(* IEC 61131-3 sources: iolistgen/tests_support/pl_stub/src/DUTs/Common, 7 files *)

(* ---- E_CmdResult.dut.st ---- *)
// Назначение: заглушка plc-process-lib 1.0.0 для проверки типов сгенерированного кода без CODESYS
//             (API.md, раздел 4.1); не библиотека — тел и внутренних переменных нет
// Автор:      kr0nsch
// Версия:     1.0.0 (выпуск библиотеки)
// Документ:   docs/GENERATORS.md, раздел «Проверка ST без CODESYS»
{attribute 'qualified_only'}
{attribute 'strict'}
TYPE E_CmdResult :
(
    None := 0,
    Accepted := 1,
    RejectedMode := 2,
    RejectedInterlock := 3,
    RejectedPermit := 4,
    RejectedInhibit := 5,
    RejectedFault := 6,
    RejectedState := 7,
    RejectedNotSupported := 8,
    RejectedCfg := 9,
    SubstExpired := 10
) INT;
END_TYPE

(* ---- E_DeviceMode.dut.st ---- *)
// Назначение: заглушка plc-process-lib 1.0.0 для проверки типов сгенерированного кода без CODESYS
//             (API.md, раздел 4.1); не библиотека — тел и внутренних переменных нет
// Автор:      kr0nsch
// Версия:     1.0.0 (выпуск библиотеки)
// Документ:   docs/GENERATORS.md, раздел «Проверка ST без CODESYS»
{attribute 'qualified_only'}
{attribute 'strict'}
TYPE E_DeviceMode :
(
    Auto := 1,
    Manual := 2,
    Local := 3,
    OutOfService := 4
) INT;
END_TYPE

(* ---- E_DeviceType.dut.st ---- *)
// Назначение: заглушка plc-process-lib 1.0.0 для проверки типов сгенерированного кода без CODESYS
//             (API.md, раздел 4.1); не библиотека — тел и внутренних переменных нет
// Автор:      kr0nsch
// Версия:     1.0.0 (выпуск библиотеки)
// Документ:   docs/GENERATORS.md, раздел «Проверка ST без CODESYS»
{attribute 'qualified_only'}
{attribute 'strict'}
TYPE E_DeviceType :
(
    None := 0,
    AnalogInput := 1,
    DigitalInput := 2,
    Motor := 3,
    MotorVfd := 4,
    Valve := 5,
    ControlValve := 6,
    Pid := 7
) INT;
END_TYPE

(* ---- E_Ne107Status.dut.st ---- *)
// Назначение: заглушка plc-process-lib 1.0.0 для проверки типов сгенерированного кода без CODESYS
//             (API.md, раздел 4.1); не библиотека — тел и внутренних переменных нет
// Автор:      kr0nsch
// Версия:     1.0.0 (выпуск библиотеки)
// Документ:   docs/GENERATORS.md, раздел «Проверка ST без CODESYS»
{attribute 'qualified_only'}
{attribute 'strict'}
TYPE E_Ne107Status :
(
    Good := 0,
    MaintenanceRequired := 1,
    OutOfSpecification := 2,
    CheckFunction := 3,
    Failure := 4
) INT;
END_TYPE

(* ---- ST_DeviceCmd.dut.st ---- *)
// Назначение: заглушка plc-process-lib 1.0.0 для проверки типов сгенерированного кода без CODESYS
//             (API.md, раздел 4.2); не библиотека — тел и внутренних переменных нет
// Автор:      kr0nsch
// Версия:     1.0.0 (выпуск библиотеки)
// Документ:   docs/GENERATORS.md, раздел «Проверка ST без CODESYS»
{attribute 'qualified_only'}
TYPE ST_DeviceCmd :
STRUCT
    xSetAuto     : BOOL;
    xSetManual   : BOOL;
    xSetOos      : BOOL;
    xReset       : BOOL;
    xAck         : BOOL;
    wAckReq      : WORD;
    wShelveReq   : WORD;
    wUnshelveReq : WORD;
END_STRUCT
END_TYPE

(* ---- ST_DeviceRetain.dut.st ---- *)
// Назначение: заглушка plc-process-lib 1.0.0 для проверки типов сгенерированного кода без CODESYS
//             (API.md, раздел 4.3); не библиотека — тел и внутренних переменных нет
// Автор:      kr0nsch
// Версия:     1.0.0 (выпуск библиотеки)
// Документ:   docs/GENERATORS.md, раздел «Проверка ST без CODESYS»
{attribute 'qualified_only'}
TYPE ST_DeviceRetain :
STRUCT
    eRemoteMode      : E_DeviceMode := E_DeviceMode.Manual;
    xOutOfService    : BOOL;
    udiOpTime_s      : UDINT;
    udiOpCount       : UDINT;
    udiOpTimeMaint_s : UDINT;
    udiOpCountMaint  : UDINT;
    // lint:allow STL007 имя массива по контракту API.md (префикс a + тип элемента)
    audiReserve      : ARRAY[0..3] OF UDINT;
END_STRUCT
END_TYPE

(* ---- ST_DeviceSts.dut.st ---- *)
// Назначение: заглушка plc-process-lib 1.0.0 для проверки типов сгенерированного кода без CODESYS
//             (API.md, раздел 4.2); не библиотека — тел и внутренних переменных нет
// Автор:      kr0nsch
// Версия:     1.0.0 (выпуск библиотеки)
// Документ:   docs/GENERATORS.md, раздел «Проверка ST без CODESYS»
{attribute 'qualified_only'}
TYPE ST_DeviceSts :
STRUCT
    wStatus     : WORD;
    wFault      : WORD;
    wWarning    : WORD;
    wCfgErr     : WORD;
    eMode       : E_DeviceMode := E_DeviceMode.Manual;
    eNe107      : E_Ne107Status := E_Ne107Status.CheckFunction;
    eCmdResult  : E_CmdResult := E_CmdResult.None;
    uiCmdSeq    : UINT;
    wAlmActive  : WORD;
    wAlmUnack   : WORD;
    wAlmShelved : WORD;
    ePrioUnack  : E_AlarmPriority := E_AlarmPriority.None;
    eDevType    : E_DeviceType := E_DeviceType.None;
    wAlmSuppressed : WORD;
END_STRUCT
END_TYPE
